Fanuc KAREL source: kt00823.compact.KL

PROGRAM KT00823
%STACKSIZE=65535
%PRIORITY=65535
%NOLOCKGROUP
VAR
R1 : REAL
R2 : REAL
OUT : REAL
BEGIN
R1=2.0
R2=3.0
R1=2.0
R2=3.0
OUT=SIN(R1)
END KT00823
